Fanuc KAREL source: kt00534.KL

PROGRAM KT00534
%STACKSIZE=65535
%PRIORITY=65535
%NOLOCKGROUP
VAR
P1 : JOINTPOS9
P2 : POSITION
OUT : POSITION
BEGIN
-- UNRESOLVED_PC line 8 opcodes [49 7E 49 60 4A] marker_code=0
END KT00534
